(*
SPDX-FileCopyrightText: © 2026 Oleksandr Tiutyk <trofimich@gmail.com>
SPDX-License-Identifier: MIT
License: https://opensource.org/license/mit
*)

(*!
<summary>Coordinates multiple child activities executing concurrently in parallel branches.</summary>
<description>
Advances all busy child activities concurrently in each execution cycle according to the configured Mode.
Under WAIT_ALL, completes when all child activities reach PASSIVE_COMPLETED. If any child halts, cancels
remaining busy children and transitions to PASSIVE_HALTED once stopped. Under WAIT_ANY, when the first child
reaches PASSIVE_COMPLETED, cancels remaining busy children and transitions to PASSIVE_COMPLETED once all
branches have safely stopped. Propagates cancellation, suspension, and resetting across all children.
</description>
*)

{attribute 'no_explicit_call' := 'do not call this function block directly'}
{attribute 'enable_dynamic_creation'}
FUNCTION_BLOCK ParallelActivity EXTENDS Activity IMPLEMENTS IParallelActivity, TOF_Core.IConfigurationSerializable
VAR_STAT
	{attribute 'hide'}
	_ClassName : STRING := __POUNAME();
END_VAR
VAR
	{attribute 'OPC.UA.DA' := '0'}
	_Children : TOF_Collections.List<0>(valueValidator := 0);

	{attribute 'OPC.UA.DA' := '0'}
	_Mode : PARALLEL_JOIN_MODE := PARALLEL_JOIN_MODE.WAIT_ALL;

	{attribute 'OPC.UA.DA' := '0'}
	_AnyBranchHalted : BOOL;

	{attribute 'OPC.UA.DA' := '0'}
	_BranchHaltReason : WSTRING(255);

	{attribute 'OPC.UA.DA' := '0'}
	_AnyBranchCompleted : BOOL;
END_VAR

(*!
<summary>Appends a child activity to be executed in parallel and returns its zero-based index.</summary>
<description>
Permitted only in PASSIVE_READY. Validates that the activity belongs to the same workflow, is not already
attached, and does not form an ancestor cycle.
The child must be unattached, including to this parent; duplicate slots are rejected before insertion.
The parent chain and owning workflow must be PASSIVE_READY. Fixed workflow association is validated.
Storage allocation precedes parent callbacks; callback exceptions may leave a partial configuration.
Child references remain borrowed and must outlive the tree. No implicit detach or ownership transfer occurs.
</description>
<param name="activity">Child activity to execute concurrently.</param>
*)
METHOD AddChildActivity : DINT
VAR_INPUT
	activity : IActivity;
END_VAR
VAR
	childParent : IWorkflowElement;
END_VAR
ValidateChildActivityAttachment(childActivity := activity, argumentName := 'activity');

childParent := activity.Parent;

IF childParent <> 0 THEN
	WorkflowExceptions.ThrowWorkflowAttachment(
		sourceNamespaceName := NamespaceName,
		sourceClassName := ClassName,
		sourcePOUName := __POUNAME(),
		sourcePosition := __POSITION(),
		message := "Child element already occupies a parent slot"
	);
END_IF

_Children.AppendGeneric(
	value := TOF_Core.GenericValueFactory.FromParts(
		genericTypeClass := TOF_Core.GENERIC_TYPE_CLASS.OBJECT,
		address := activity.SelfAddress,
		size := activity.SelfSize,
		memoryManagementBehavior := TOF_Core.GENERIC_MEMORY_MANAGEMENT_BEHAVIOR.STORE_ORIGINAL_REFERENCE_AND_NOT_OWNS_MEMORY
	),
	index => AddChildActivity
);

activity.ParentActivity := THIS^;
END_METHOD

(*!
<summary>Returns the number of child activities registered for parallel execution.</summary>
*)
{attribute 'monitoring' := 'call'}
PROPERTY ChildCount : DINT
GET
ChildCount := _Children.Length;
END_GET
END_PROPERTY

(*!
<summary>Borrows the initialized class name used in diagnostics.</summary>
<description>
Returns initialized metadata storage without allocation. Callers must not modify the returned string.
Derived function blocks must use distinct initialized static storage when overriding this metadata.
</description>
*)
{attribute 'monitoring' := 'call'}
PROPERTY ClassName : REFERENCE TO STRING
GET
ClassName REF= _ClassName;
END_GET
END_PROPERTY

(*!
<summary>Returns the child activity at the specified zero-based index, or 0 if the index is out of bounds.</summary>
<param name="index">Zero-based index of the child activity.</param>
*)
METHOD GetChildActivity : IActivity
VAR_INPUT
	index : DINT;
END_VAR
IF index >= TOF_Core.SignedInt32.ZERO AND_THEN index < _Children.Length THEN
	__QUERYINTERFACE(_Children.Get(index := index).AsObject(), GetChildActivity);
END_IF
END_METHOD

(*!
<summary>Gets or sets the join completion mode (WAIT_ALL or WAIT_ANY).</summary>
<description>
Can only be modified while the activity is in PASSIVE_READY.
</description>
*)
{attribute 'monitoring' := 'call'}
PROPERTY Mode : PARALLEL_JOIN_MODE
GET
Mode := _Mode;
END_GET
SET
IF State <> WORKFLOW_ELEMENT_STATE.PASSIVE_READY THEN
	WorkflowExceptions.ThrowWorkflowConfiguration(
		sourceNamespaceName := NamespaceName,
		sourceClassName := ClassName,
		sourcePOUName := __POUNAME(),
		sourcePosition := __POSITION(),
		message := "Cannot modify parallel join mode outside PASSIVE_READY"
	);
END_IF

_Mode := Mode;
END_SET
END_PROPERTY

(*!
<summary>Borrows the compiler-initialized library namespace.</summary>
<description>
Borrows storage from the live internal namespace provider. Reacquire references after application
reinitialization or relocation. Treat the reference as read-only; no ownership or synchronization is provided.
</description>
*)
{attribute 'monitoring' := 'call'}
PROPERTY NamespaceName : REFERENCE TO STRING
GET
NamespaceName REF= CurrentNamespace.Name;
END_GET
END_PROPERTY

(*!
<summary>Cancels all active child activities when this parallel activity transitions to PASSIVE_FAILED.</summary>
<description>
Attempts cancellation of each busy child independently under the no-throw hook contract. It does not wait
for child stopping or release. Child cancellation failures preserve the parent failure; OnResetting or the
explicit resource owner must finish recovery before affected resources are reused.
</description>
<param name="exception">Caught exception that caused the failure.</param>
*)
METHOD PROTECTED OnFail
VAR_INPUT
	exception : TOF_Core.IException;
END_VAR
VAR
	i : DINT;
	child : IActivity;
END_VAR
FOR i := 0 TO _Children.Length - 1 DO
	child := GetChildActivity(index := i);

	IF child <> 0 AND_THEN child.Busy THEN
		__TRY
			child.RequestCancel(reason := "Parent parallel activity failed");
		__CATCH
		__ENDTRY
	END_IF
END_FOR
END_METHOD

(*!
<summary>Drives resetting of all non-ready child activities back to PASSIVE_READY.</summary>
<param name="startResetting">TRUE on the initial call from RequestReset.</param>
*)
METHOD PROTECTED OnResetting : ACTIVITY_RESETTING_STATE
VAR_INPUT
	startResetting : BOOL;
END_VAR
VAR
	i : DINT;
	child : IActivity;
	allReset : BOOL;
END_VAR
IF _Children.Length = TOF_Core.SignedInt32.ZERO THEN
	_AnyBranchHalted := FALSE;
	_BranchHaltReason := "";
	_AnyBranchCompleted := FALSE;
	OnResetting := ACTIVITY_RESETTING_STATE.WORK_RESET;
	RETURN;
END_IF

allReset := TRUE;

FOR i := 0 TO _Children.Length - 1 DO
	child := GetChildActivity(index := i);

	IF child <> 0 AND_THEN child.State <> WORKFLOW_ELEMENT_STATE.PASSIVE_READY THEN
		IF ResetChildActivity(childActivity := child) = ACTIVITY_RESETTING_STATE.WORK_IN_PROGRESS THEN
			allReset := FALSE;
		END_IF
	END_IF
END_FOR

IF allReset THEN
	_AnyBranchHalted := FALSE;
	_BranchHaltReason := "";
	_AnyBranchCompleted := FALSE;
	OnResetting := ACTIVITY_RESETTING_STATE.WORK_RESET;
ELSE
	OnResetting := ACTIVITY_RESETTING_STATE.WORK_IN_PROGRESS;
END_IF
END_METHOD

(*!
<summary>Advances all busy child activities concurrently and evaluates parallel join completion.</summary>
<param name="startRunning">TRUE on the initial call of a fresh start from PASSIVE_READY.</param>
<param name="startResuming">TRUE on the initial call when resuming from PASSIVE_SUSPENDED.</param>
<param name="haltReason">Receives the diagnostic reason if a child activity halts.</param>
*)
METHOD PROTECTED OnRunning : ACTIVITY_RUNNING_STATE
VAR_INPUT
	startRunning : BOOL;
	startResuming : BOOL;
END_VAR
VAR_OUTPUT
	haltReason : WSTRING(255);
END_VAR
VAR
	i : DINT;
	child : IActivity;
	allCompleted : BOOL;
	anyBusy : BOOL;
END_VAR
IF _Children.Length = TOF_Core.SignedInt32.ZERO THEN
	_AnyBranchHalted := FALSE;
	_BranchHaltReason := "";
	_AnyBranchCompleted := FALSE;
	OnRunning := ACTIVITY_RUNNING_STATE.WORK_COMPLETED;
	RETURN;
END_IF

IF startRunning THEN
	_AnyBranchHalted := FALSE;
	_BranchHaltReason := "";
	_AnyBranchCompleted := FALSE;

	FOR i := 0 TO _Children.Length - 1 DO
		child := GetChildActivity(index := i);

		IF child <> 0 THEN
			child.RequestStart();
		END_IF
	END_FOR
ELSIF startResuming THEN
	FOR i := 0 TO _Children.Length - 1 DO
		child := GetChildActivity(index := i);

		IF child <> 0 AND_THEN child.State = WORKFLOW_ELEMENT_STATE.PASSIVE_SUSPENDED THEN
			child.RequestStart();
		END_IF
	END_FOR
ELSE
	FOR i := 0 TO _Children.Length - 1 DO
		child := GetChildActivity(index := i);

		IF child <> 0 AND_THEN child.Busy THEN
			child.Execute();
		END_IF
	END_FOR
END_IF

allCompleted := TRUE;
anyBusy := FALSE;

FOR i := 0 TO _Children.Length - 1 DO
	child := GetChildActivity(index := i);

	IF child <> 0 THEN
		IF child.Busy THEN
			anyBusy := TRUE;
			allCompleted := FALSE;
		ELSIF child.State = WORKFLOW_ELEMENT_STATE.PASSIVE_COMPLETED THEN
			_AnyBranchCompleted := TRUE;
		ELSIF child.State = WORKFLOW_ELEMENT_STATE.PASSIVE_HALTED THEN
			allCompleted := FALSE;

			IF NOT _AnyBranchHalted THEN
				_AnyBranchHalted := TRUE;
				_BranchHaltReason := child.HaltReason;
			END_IF
		ELSE
			allCompleted := FALSE;
		END_IF
	END_IF
END_FOR

IF _AnyBranchHalted THEN
	IF anyBusy THEN
		FOR i := 0 TO _Children.Length - 1 DO
			child := GetChildActivity(index := i);

			IF child <> 0 AND_THEN child.Busy AND_THEN child.State <> WORKFLOW_ELEMENT_STATE.ACTIVE_CANCELLING THEN
				child.RequestCancel(reason := "Parallel sibling branch halted");
			END_IF
		END_FOR

		OnRunning := ACTIVITY_RUNNING_STATE.WORK_IN_PROGRESS;
	ELSE
		haltReason := _BranchHaltReason;
		OnRunning := ACTIVITY_RUNNING_STATE.WORK_HALTED;
	END_IF

	RETURN;
END_IF

IF _Mode = PARALLEL_JOIN_MODE.WAIT_ANY AND_THEN _AnyBranchCompleted THEN
	IF anyBusy THEN
		FOR i := 0 TO _Children.Length - 1 DO
			child := GetChildActivity(index := i);

			IF child <> 0 AND_THEN child.Busy AND_THEN child.State <> WORKFLOW_ELEMENT_STATE.ACTIVE_CANCELLING THEN
				child.RequestCancel(reason := "Parallel branch completed (WAIT_ANY)");
			END_IF
		END_FOR

		OnRunning := ACTIVITY_RUNNING_STATE.WORK_IN_PROGRESS;
	ELSE
		OnRunning := ACTIVITY_RUNNING_STATE.WORK_COMPLETED;
	END_IF

	RETURN;
END_IF

IF allCompleted THEN
	OnRunning := ACTIVITY_RUNNING_STATE.WORK_COMPLETED;
ELSE
	OnRunning := ACTIVITY_RUNNING_STATE.WORK_IN_PROGRESS;
END_IF
END_METHOD

(*!
<summary>Stops all active child activities cooperatively and waits for them to reach a passive state.</summary>
<param name="startCancelling">TRUE on the initial call from RequestCancel.</param>
<param name="startSuspending">TRUE on the initial call from RequestSuspend.</param>
<param name="haltReason">Receives the diagnostic reason if a child activity halts while stopping.</param>
*)
METHOD PROTECTED OnStopping : ACTIVITY_STOPPING_STATE
VAR_INPUT
	startCancelling : BOOL;
	startSuspending : BOOL;
END_VAR
VAR_OUTPUT
	haltReason : WSTRING(255);
END_VAR
VAR
	i : DINT;
	child : IActivity;
	anyBusy : BOOL;
	anyHalted : BOOL;
	allCompleted : BOOL;
END_VAR
IF _Children.Length = TOF_Core.SignedInt32.ZERO THEN
	OnStopping := ACTIVITY_STOPPING_STATE.WORK_STOPPED;
	RETURN;
END_IF

IF startCancelling THEN
	FOR i := 0 TO _Children.Length - 1 DO
		child := GetChildActivity(index := i);

		IF child <> 0 THEN
			IF child.Busy THEN
				child.RequestCancel(reason := _CancelReason);
			ELSIF child.State = WORKFLOW_ELEMENT_STATE.PASSIVE_SUSPENDED THEN
				child.RequestCancel(reason := _CancelReason);
			END_IF
		END_IF
	END_FOR
ELSIF startSuspending THEN
	FOR i := 0 TO _Children.Length - 1 DO
		child := GetChildActivity(index := i);

		IF child <> 0 AND_THEN child.Busy THEN
			child.RequestSuspend();
		END_IF
	END_FOR
ELSE
	FOR i := 0 TO _Children.Length - 1 DO
		child := GetChildActivity(index := i);

		IF child <> 0 AND_THEN child.Busy THEN
			child.Execute();
		END_IF
	END_FOR
END_IF

anyBusy := FALSE;
anyHalted := FALSE;
allCompleted := TRUE;

FOR i := 0 TO _Children.Length - 1 DO
	child := GetChildActivity(index := i);

	IF child <> 0 THEN
		IF child.Busy THEN
			anyBusy := TRUE;
			allCompleted := FALSE;
		ELSIF child.State = WORKFLOW_ELEMENT_STATE.PASSIVE_HALTED THEN
			allCompleted := FALSE;

			IF NOT anyHalted THEN
				anyHalted := TRUE;

				IF _BranchHaltReason = "" THEN
					_BranchHaltReason := child.HaltReason;
				END_IF
			END_IF
		ELSIF child.State <> WORKFLOW_ELEMENT_STATE.PASSIVE_COMPLETED THEN
			allCompleted := FALSE;
		END_IF
	END_IF
END_FOR

IF anyBusy THEN
	OnStopping := ACTIVITY_STOPPING_STATE.WORK_IN_PROGRESS;
	RETURN;
END_IF

IF anyHalted OR_ELSE _AnyBranchHalted THEN
	haltReason := _BranchHaltReason;
	OnStopping := ACTIVITY_STOPPING_STATE.WORK_HALTED;
ELSIF allCompleted THEN
	OnStopping := ACTIVITY_STOPPING_STATE.WORK_COMPLETED;
ELSE
	OnStopping := ACTIVITY_STOPPING_STATE.WORK_STOPPED;
END_IF
END_METHOD

(*!
<summary>Advances resetting of a child activity toward PASSIVE_READY by one step.</summary>
<description>
Returns WORK_RESET immediately when childActivity is 0 or already in PASSIVE_READY. If the child was left in
PASSIVE_SUSPENDED or ACTIVE_CANCELLING, drives cancellation to PASSIVE_CANCELLED before invoking RequestReset.
In ACTIVE_RESETTING, advances the child via Execute; in finished passive states, invokes RequestReset.
</description>
<param name="childActivity">Child activity to reset, or 0.</param>
*)
METHOD PROTECTED ResetChildActivity : ACTIVITY_RESETTING_STATE
VAR_INPUT
	childActivity : IActivity;
END_VAR
ResetChildActivity := WorkflowElementHelper.ResetChildActivity(
	childActivity := childActivity,
	cancelReason := "Parent parallel activity resetting",
	sourceClassName := ClassName,
	sourcePOUName := __POUNAME()
);
END_METHOD

(*!
<summary>Reports the size of this concrete function block instance in bytes.</summary>
<description>
Reports the instance layout rather than dynamic allocations owned by its fields. A derived function block
with a different layout must override this property; the value does not grant disposal rights.
</description>
*)
{attribute 'monitoring' := 'call'}
PROPERTY SelfSize : ULINT
GET
SelfSize := XSIZEOF(THIS^);
END_GET
END_PROPERTY

(*!
<summary>
Verifies that a candidate child activity can be attached to this parallel composite without cycles or
conflicts.
</summary>
<description>
Delegates to Workflows.ValidateElementAttachment for readiness, cycles, existing parent, root exclusion and
fixed workflow association. Reusing the same link during Configure is allowed; append methods must reject
occupied slots separately. No topology or ownership mutation is performed.
</description>
<param name="childActivity">Candidate child activity to validate.</param>
<param name="argumentName">Parameter name for diagnostic reporting.</param>
*)
METHOD PROTECTED ValidateChildActivityAttachment
VAR_INPUT
	childActivity : IActivity;
	argumentName : STRING(255);
END_VAR
WorkflowElementHelper.ValidateChildActivityAttachment(
	parent := THIS^,
	childActivity := childActivity,
	argumentName := argumentName,
	sourceClassName := ClassName,
	sourcePOUName := __POUNAME()
);
END_METHOD

(*!
<summary>Writes the configuration fields for this object.</summary>
<description>Borrows the writer for this call. A failure invalidates the current output document.</description>
*)
METHOD Serialize
VAR_INPUT
	writer : TOF_Core.IConfigurationWriter;
END_VAR
VAR
	mode : DINT;
	i : DINT;
END_VAR
Workflows.WriteConfigurationHeader(writer := writer, source := THIS^, displayName := Name, scope := THIS^);
mode := TO_DINT(_Mode);
writer.WriteValue(
	name := 'mode',
	valueType := TOF_Core.CONFIGURATION_VALUE_TYPE.TYPE_DINT,
	data := ADR(mode),
	size := SIZEOF(mode)
);
writer.BeginArray(name := 'children');

FOR i := 0 TO _Children.Length - 1 DO
	Workflows.WriteConfigurationObject(writer := writer, name := '', source := _Children.Get(index := i).AsObject());
END_FOR

writer.EndArray();
END_METHOD

(*!
<summary>Restores this fresh instance from its configuration object.</summary>
<description>
The reader, document node and deserialization context are borrowed for this call.
On failure discard the partial instance.
</description>
<param name="reader">Active configuration reader.</param>
<param name="node">Object node to read fields from.</param>
<param name="context">Active configuration deserialization context providing workflow reconstruction services.</param>
*)
METHOD Deserialize
VAR_INPUT
	reader : TOF_Core.IConfigurationReader;
	node : TOF_Core.CONFIGURATION_NODE;
	context : TOF_Core.IConfigurationDeserializationContext;
END_VAR
VAR
	loader : IWorkflowLoader;
	items : TOF_Core.CONFIGURATION_NODE;
	count : DINT;
	i : DINT;
	code : DINT;
END_VAR
loader := WorkflowConfigurationSerializer.ResolveWorkflowLoader(context := context);
Workflows.ReadConfigurationHeader(reader := reader, node := node, target := THIS^, scope := THIS^);

reader.ReadValue(
	node := reader.GetField(node := node, name := 'mode'),
	valueType := TOF_Core.CONFIGURATION_VALUE_TYPE.TYPE_DINT,
	data := ADR(code),
	size := SIZEOF(code)
);

CASE code OF
	0:
		Mode := PARALLEL_JOIN_MODE.WAIT_ALL;
	1:
		Mode := PARALLEL_JOIN_MODE.WAIT_ANY;
ELSE
	WorkflowExceptions.ThrowWorkflowConfiguration(
		sourceNamespaceName := NamespaceName,
		sourceClassName := ClassName,
		sourcePOUName := __POUNAME(),
		sourcePosition := __POSITION(),
		message := "Unknown mode value"
	);
END_CASE

items := reader.GetField(node := node, name := 'children');
count := TO_DINT(reader.GetArraySize(node := items));

FOR i := 0 TO count - 1 DO
	AddChildActivity(
		activity := Workflows.ReadActivity(loader := loader, node := reader.GetItem(node := items, index := TO_UDINT(i)))
	);
END_FOR
END_METHOD

END_FUNCTION_BLOCK

(* stored: Version 1.1.0.1
   POU ParallelActivity: Id {6c5ddb07-2877-413c-a1a1-f1e269fb6def}, SpecialFunc None
   Folder Overriden methods: Id {885741b9-d520-4a51-9f57-e60d9237c02b}
   Folder Service methods: Id {7baed18b-ddb6-4a91-b4cc-1407e3826a3f}
   Method AddChildActivity: Id {0292ec90-8c9b-4d75-b95c-7d712d77dd0f}
   Property ChildCount: Id {f1d507c7-8363-4045-a8d3-b5afa6acf345}
   Get Get: Id {c3962e91-9a15-4b7f-a47a-e846d6b53c5b}
   Property ClassName: Id {f108a989-028d-405d-87cf-71f0f548a4d6}
   Get Get: Id {e13e85c6-7fb6-49a2-bb4c-1ac98668a3d5}
   Method GetChildActivity: Id {2954fc95-78c9-4fde-a38b-2c20fa1f2471}
   Property Mode: Id {58a2c073-b79d-497c-818c-5b08eed0876e}
   Get Get: Id {1924c67c-4f95-4132-b4d7-95ec46fb3d61}
   Set Set: Id {7bec509a-a3f2-481b-a9f3-cf6a6bff1473}
   Property NamespaceName: Id {b01d14a2-cf3c-4554-83c0-3da70ecb2e96}
   Get Get: Id {e65dc63c-0d39-4335-b979-44071d360f90}
   Method OnFail: Id {0d7481d5-e08f-41df-bce5-678c7c1a7ebe}
   Method OnResetting: Id {59a532c0-886c-4108-9fd7-fbea264997ee}
   Method OnRunning: Id {83a490b1-f30e-48d1-81a8-4c4cf4e6def3}
   Method OnStopping: Id {e5406289-8349-40c6-ac4a-67e538744cfa}
   Method ResetChildActivity: Id {92256385-9c2d-41ca-b895-4719a423bc33}
   Property SelfSize: Id {a91f65a8-cf85-4b20-a318-aec1e1d0f781}
   Get Get: Id {63d24e9a-fedc-40ac-9fcc-d98ab14927ae}
   Method ValidateChildActivityAttachment: Id {d9ebf347-b252-46ff-91b8-1ef334536ad6}
   Method Serialize: Id {b69ec900-bb90-4c4d-a34f-f88bc5fefb2f}
   Method Deserialize: Id {d8b67d7f-18d1-45ab-87bf-7bb9b2b8df03} *)
